(* IEC 61131-3 sources: jwplc-sim/tests/openplc/blink-alias/pous/programs, 1 file *)

(* ---- main.st ---- *)
PROGRAM main
  VAR
    Q0_0_OUT AT Out0 : BOOL;
    Q0_1_OUT AT Out1 : BOOL;
    I0_0_IN AT Int0 : BOOL;
    T1 : TON;
    T2 : TON;
  END_VAR

  T1(IN := NOT T2.Q, PT := T#500ms);
  T2(IN := T1.Q, PT := T#500ms);
  Q0_0_OUT := T1.Q;
  Q0_1_OUT := I0_0_IN;

END_PROGRAM
